PROGRAM MAIN
VAR
	Machine : UM_Tutorial := (Description := ' Tutorial Project ',
							UseGenericVISU := TRUE);
	DownloadBit : BOOL := TRUE;
END_VAR

TT_GIO.Safety(Reset_Trigger := Machine.PbReset.Actuate);
TT_GIO.Safety.In.EStop_OK := TRUE;
TT_GIO.Safety.In.EStop_STO := TRUE;

Machine(SafetyBlock := TT_GIO.Safety);

END_PROGRAM

(* stored: Version 1.1.0.1, ProductVersion 3.1.4024.12
   POU MAIN: Id {81a9f757-7db3-43f0-a54f-2190313d9fed}, SpecialFunc None *)
